// #272: an elevation error during a slew. In the scan of the error only the elevation is disabled and the shared brake is
// closed (no drive holds it); azimuth and derotator stay enabled and get their MC_Stop at the fast-stop dynamics of stMotion
// (bAxisErrorRamp), the hydraulics stay on. After the stop has settled the emergency park parks in place: all axes disabled,
// brake closed, covers closed, hydraulics off, the stop dynamics back at the NC parameters (0.0). Until 0.23.x all three axes
// were disabled in the scan of the error and the brake alone stopped the azimuth.
// #277: the azimuth drive (the NC enable behind the HalfBROT brake gate, fbAxis.Ready in the mock) stays on during the ramp
// although the shared brake is closed (HalfBROT FB_BrakeCloseHold); without the hold the gate dropped it in the next scan.
METHOD PRIVATE Elevation_Error_During_A_Slew_Fast_Stops_The_Healthy_Axes
VAR_INST
	pRig		: POINTER TO FB_MonetRig;	// created with __NEW in this test's turn, freed in the scan it finished in
	rig			: REFERENCE TO FB_MonetRig;
	stCfg		: BROTLib.ST_MotionConfig;
	nStep		: INT;
	nCycles		: UINT;
	sTest		: STRING(80);
	nAz0		: UINT;
	nDr0		: UINT;
	nDisable0	: UINT;
	bSeenError	: BOOL;
	bSawRamp	: BOOL;
	bAzDriveLost	: BOOL;	// #277: a ramp scan with the azimuth wanted enabled but its drive off
END_VAR
TEST('Elevation_Error_During_A_Slew_Fast_Stops_The_Healthy_Axes');
sTest := 'Elevation_Error_During_A_Slew_Fast_Stops_The_Healthy_Axes: ';
IF nStep >= 90 THEN
	RETURN;
END_IF
IF nCur <> 22 THEN	// not this test's turn yet (TEST() above is called in every scan, TcUnit needs that)
	RETURN;
END_IF
IF pRig = 0 THEN
	pRig := __NEW(FB_MonetRig);
	IF pRig = 0 THEN
		AssertTrue(Condition := FALSE, Message := 'no router memory for the rig');
		F_Note(bFailed := TRUE, sText := CONCAT(sTest, 'no router memory for the rig'));
		nStep := 99;
		nCur := nCur + 1;
		TEST_FINISHED();
		RETURN;
	END_IF
	rig REF= pRig^;
END_IF
IF nStep = 0 AND nCycles = 0 THEN
	stCfg.fAzimuthFastStopDeceleration := 10.0;
	stCfg.fAzimuthFastStopJerk := 30.0;
	stCfg.fElevationFastStopDeceleration := 9.0;
	stCfg.fElevationFastStopJerk := 27.0;
	stCfg.fDerotatorFastStopDeceleration := 20.0;
	stCfg.fDerotatorFastStopJerk := 60.0;
	rig.SetMotion(stValue := stCfg);
END_IF
rig.Scan();
nCycles := nCycles + 1;
CASE nStep OF
0:	// wait for the clock, then power on
	IF rig.ClockValid THEN
		rig.fbTel.Init();
		nStep := 10;
		nCycles := 0;
	ELSIF nCycles > 2000 THEN
		AssertTrue(Condition := FALSE, Message := 'the astronomical clock never became valid');
		F_Note(bFailed := TRUE, sText := CONCAT(sTest, 'the astronomical clock never became valid'));
		nStep := 99;
		TEST_FINISHED();
	END_IF
10:	// online: slew
	IF rig.Online THEN
		rig.fbTel.Slew(fAzimuth := 180.0, fAltitude := 45.0);
		nStep := 20;
		nCycles := 0;
	ELSIF nCycles > 1500 THEN
		AssertTrue(Condition := FALSE, Message := 'the mock telescope did not reach READY_STATE 1.0');
		F_Note(bFailed := TRUE, sText := CONCAT(sTest, 'the mock telescope did not reach READY_STATE 1.0'));
		nStep := 99;
		TEST_FINISHED();
	END_IF
20:	// the slew moves all three axes: the elevation reports an error
	IF rig.fbElev.MoveAxis AND rig.fbAzim.MoveAxis AND rig.fbDero.MoveAxis AND nCycles >= 3 THEN
		nAz0 := rig.fbAzim.nStopEdges;
		nDr0 := rig.fbDero.nStopEdges;
		nDisable0 := rig.fbBrakeHyd.nDisableCalls;
		rig.InjectElevationError(16#4550);
		nStep := 30;
		nCycles := 0;
	ELSIF nCycles > 300 THEN
		AssertTrue(Condition := FALSE, Message := 'the slew did not start the axis moves');
		F_Note(bFailed := TRUE, sText := CONCAT(sTest, 'the slew did not start the axis moves'));
		nStep := 99;
		TEST_FINISHED();
	END_IF
30:
	bSawRamp := bSawRamp OR rig.fbTel.bAxisErrorRamp;
	// the drive off while the azimuth still moves or stops (the mock core keeps moving without its enable)
	IF rig.fbTel.bAxisErrorRamp AND rig.fbAzim.bEnable AND NOT rig.fbAzim.fbAxis.Ready AND NOT rig.fbAzim.fbAxis.StandStill THEN
		bAzDriveLost := TRUE;
	END_IF
	IF rig.fbTel.bError AND NOT bSeenError THEN	// the scan that saw the error
		bSeenError := TRUE;
		AssertTrue(Condition := rig.fbTel.bAxisErrorRamp AND rig.fbTel.bStopActive, Message := 'the error starts the ramp (bStop)');
		F_Note(bFailed := NOT (rig.fbTel.bAxisErrorRamp AND rig.fbTel.bStopActive), sText := CONCAT(sTest, 'the error starts the ramp (bStop)'));
		AssertFalse(Condition := rig.fbElev.bEnable, Message := 'the faulty elevation is disabled');
		F_Note(bFailed := (rig.fbElev.bEnable), sText := CONCAT(sTest, 'the faulty elevation is disabled'));
		AssertTrue(Condition := rig.fbAzim.bEnable AND rig.fbDero.bEnable, Message := 'azimuth and derotator stay enabled for their stop');
		F_Note(bFailed := NOT (rig.fbAzim.bEnable AND rig.fbDero.bEnable), sText := CONCAT(sTest, 'azimuth and derotator stay enabled for their stop'));
		AssertFalse(Condition := rig.fbBrakeHyd.BrakeOpen, Message := 'the shared brake is closed at once');
		F_Note(bFailed := (rig.fbBrakeHyd.BrakeOpen), sText := CONCAT(sTest, 'the shared brake is closed at once'));
		AssertTrue(Condition := rig.fbBrakeHyd.nDisableCalls = nDisable0, Message := 'the hydraulics stay on');
		F_Note(bFailed := NOT (rig.fbBrakeHyd.nDisableCalls = nDisable0), sText := CONCAT(sTest, 'the hydraulics stay on'));
		AssertTrue(Condition := rig.fbAzim.fbAxis.StopDeceleration = 10.0 AND rig.fbAzim.fbAxis.StopJerk = 30.0, Message := 'the azimuth stops at its fast-stop dynamics');
		F_Note(bFailed := NOT (rig.fbAzim.fbAxis.StopDeceleration = 10.0 AND rig.fbAzim.fbAxis.StopJerk = 30.0), sText := CONCAT(sTest, 'the azimuth stops at its fast-stop dynamics'));
		AssertTrue(Condition := rig.fbDero.fbAxis.StopDeceleration = 20.0 AND rig.fbDero.fbAxis.StopJerk = 60.0, Message := 'the derotator stops at its fast-stop dynamics');
		F_Note(bFailed := NOT (rig.fbDero.fbAxis.StopDeceleration = 20.0 AND rig.fbDero.fbAxis.StopJerk = 60.0), sText := CONCAT(sTest, 'the derotator stops at its fast-stop dynamics'));
	END_IF
	IF rig.fbTel.bIsParked AND nCycles > 5 THEN
		AssertTrue(Condition := bSawRamp, Message := 'the ramp ran');
		F_Note(bFailed := NOT (bSawRamp), sText := CONCAT(sTest, 'the ramp ran'));
		AssertFalse(Condition := bAzDriveLost, Message := 'the azimuth drive stays on for its stop with the brake closed');
		F_Note(bFailed := bAzDriveLost, sText := CONCAT(sTest, 'the azimuth drive stays on for its stop with the brake closed'));
		AssertTrue(Condition := rig.fbAzim.nStopEdges > nAz0 AND rig.fbDero.nStopEdges > nDr0, Message := 'azimuth and derotator were sent their MC_Stop');
		F_Note(bFailed := NOT (rig.fbAzim.nStopEdges > nAz0 AND rig.fbDero.nStopEdges > nDr0), sText := CONCAT(sTest, 'azimuth and derotator were sent their MC_Stop'));
		AssertTrue(Condition := rig.fbTel.bParkedInPlace AND NOT rig.fbTel.bParkActive AND NOT rig.fbTel.bAxisErrorRamp, Message := 'the park ended in place, the ramp is over');
		F_Note(bFailed := NOT (rig.fbTel.bParkedInPlace AND NOT rig.fbTel.bParkActive AND NOT rig.fbTel.bAxisErrorRamp), sText := CONCAT(sTest, 'the park ended in place, the ramp is over'));
		AssertFalse(Condition := rig.fbElev.bEnable OR rig.fbAzim.bEnable OR rig.fbDero.bEnable, Message := 'all three axes are disabled');
		F_Note(bFailed := (rig.fbElev.bEnable OR rig.fbAzim.bEnable OR rig.fbDero.bEnable), sText := CONCAT(sTest, 'all three axes are disabled'));
		AssertFalse(Condition := rig.fbBrakeHyd.BrakeOpen, Message := 'the brake is closed');
		F_Note(bFailed := (rig.fbBrakeHyd.BrakeOpen), sText := CONCAT(sTest, 'the brake is closed'));
		AssertTrue(Condition := rig.fbCovers.bClosed AND rig.fbBrakeHyd.nDisableCalls > nDisable0, Message := 'covers closed, hydraulics off');
		F_Note(bFailed := NOT (rig.fbCovers.bClosed AND rig.fbBrakeHyd.nDisableCalls > nDisable0), sText := CONCAT(sTest, 'covers closed, hydraulics off'));
		AssertTrue(Condition := rig.fbAzim.fbAxis.StopDeceleration = 0.0 AND rig.fbAzim.fbAxis.StopJerk = 0.0 AND
			rig.fbDero.fbAxis.StopDeceleration = 0.0 AND rig.fbElev.fbAxis.StopDeceleration = 0.0, Message := 'the stop dynamics are back at the NC parameters');
		F_Note(bFailed := NOT (rig.fbAzim.fbAxis.StopDeceleration = 0.0 AND rig.fbAzim.fbAxis.StopJerk = 0.0 AND
			rig.fbDero.fbAxis.StopDeceleration = 0.0 AND rig.fbElev.fbAxis.StopDeceleration = 0.0), sText := CONCAT(sTest, 'the stop dynamics are back at the NC parameters'));
		AssertTrue(Condition := rig.fbTel.bError AND rig.fbTel.ReadyState = -1.0, Message := 'the error stays, READY_STATE -1.0');
		F_Note(bFailed := NOT (rig.fbTel.bError AND rig.fbTel.ReadyState = -1.0), sText := CONCAT(sTest, 'the error stays, READY_STATE -1.0'));
		nStep := 99;
		TEST_FINISHED();
	ELSIF nCycles > 1000 THEN
		AssertTrue(Condition := FALSE, Message := 'the telescope did not park after the ramp');
		F_Note(bFailed := TRUE, sText := CONCAT(sTest, 'the telescope did not park after the ramp'));
		nStep := 99;
		TEST_FINISHED();
	END_IF
END_CASE
IF nStep >= 90 AND pRig <> 0 THEN	// finished in this scan: free the rig, the next test starts in the next scan
	__DELETE(pRig);
	pRig := 0;
	nCur := nCur + 1;
END_IF
END_METHOD

// #272: an azimuth error during a slew. The faulty azimuth has no drive, so the shared brake is closed in the scan of the error
// (until 0.23.x the emergency park closed it in that scan; the park now waits behind the ramp) and held closed: the enabled
// elevation requests the opening in every scan. Elevation and derotator stay enabled and get their MC_Stop; then the park parks
// in place. #277: the elevation drive stays on for its stop although the brake is closed (HalfBROT FB_BrakeCloseHold).
METHOD PRIVATE Azimuth_Error_During_A_Slew_Closes_The_Brake_At_Once
VAR_INST
	pRig		: POINTER TO FB_MonetRig;	// created with __NEW in this test's turn, freed in the scan it finished in
	rig			: REFERENCE TO FB_MonetRig;
	nStep		: INT;
	nCycles		: UINT;
	sTest		: STRING(80);
	nEl0		: UINT;
	nDisable0	: UINT;
	bSeenError	: BOOL;
	bReopened	: BOOL;	// the brake was open again in a later scan of the ramp (the enabled elevation requests the opening in every scan)
	bElDriveLost	: BOOL;	// #277: a ramp scan with the elevation wanted enabled but its drive off while it still moves
END_VAR
TEST('Azimuth_Error_During_A_Slew_Closes_The_Brake_At_Once');
sTest := 'Azimuth_Error_During_A_Slew_Closes_The_Brake_At_Once: ';
IF nStep >= 90 THEN
	RETURN;
END_IF
IF nCur <> 23 THEN	// not this test's turn yet (TEST() above is called in every scan, TcUnit needs that)
	RETURN;
END_IF
IF pRig = 0 THEN
	pRig := __NEW(FB_MonetRig);
	IF pRig = 0 THEN
		AssertTrue(Condition := FALSE, Message := 'no router memory for the rig');
		F_Note(bFailed := TRUE, sText := CONCAT(sTest, 'no router memory for the rig'));
		nStep := 99;
		nCur := nCur + 1;
		TEST_FINISHED();
		RETURN;
	END_IF
	rig REF= pRig^;
END_IF
rig.Scan();
nCycles := nCycles + 1;
CASE nStep OF
0:	// wait for the clock, then power on
	IF rig.ClockValid THEN
		rig.fbTel.Init();
		nStep := 10;
		nCycles := 0;
	ELSIF nCycles > 2000 THEN
		AssertTrue(Condition := FALSE, Message := 'the astronomical clock never became valid');
		F_Note(bFailed := TRUE, sText := CONCAT(sTest, 'the astronomical clock never became valid'));
		nStep := 99;
		TEST_FINISHED();
	END_IF
10:	// online: slew
	IF rig.Online THEN
		rig.fbTel.Slew(fAzimuth := 180.0, fAltitude := 45.0);
		nStep := 20;
		nCycles := 0;
	ELSIF nCycles > 1500 THEN
		AssertTrue(Condition := FALSE, Message := 'the mock telescope did not reach READY_STATE 1.0');
		F_Note(bFailed := TRUE, sText := CONCAT(sTest, 'the mock telescope did not reach READY_STATE 1.0'));
		nStep := 99;
		TEST_FINISHED();
	END_IF
20:	// the slew moves all three axes: the azimuth reports an error
	IF rig.fbElev.MoveAxis AND rig.fbAzim.MoveAxis AND rig.fbDero.MoveAxis AND nCycles >= 3 THEN
		nEl0 := rig.fbElev.nStopEdges;
		nDisable0 := rig.fbBrakeHyd.nDisableCalls;
		rig.InjectAzimuthError(16#4550);
		nStep := 30;
		nCycles := 0;
	ELSIF nCycles > 300 THEN
		AssertTrue(Condition := FALSE, Message := 'the slew did not start the axis moves');
		F_Note(bFailed := TRUE, sText := CONCAT(sTest, 'the slew did not start the axis moves'));
		nStep := 99;
		TEST_FINISHED();
	END_IF
30:
	IF rig.fbTel.bAxisErrorRamp AND rig.fbElev.bEnable AND NOT rig.fbElev.fbAxis.Ready AND NOT rig.fbElev.fbAxis.StandStill THEN
		bElDriveLost := TRUE;
	END_IF
	IF rig.fbTel.bError AND NOT bSeenError THEN	// the scan that saw the error
		bSeenError := TRUE;
		AssertTrue(Condition := rig.fbTel.bAxisErrorRamp, Message := 'the error starts the ramp');
		F_Note(bFailed := NOT (rig.fbTel.bAxisErrorRamp), sText := CONCAT(sTest, 'the error starts the ramp'));
		AssertFalse(Condition := rig.fbAzim.bEnable, Message := 'the faulty azimuth is disabled');
		F_Note(bFailed := (rig.fbAzim.bEnable), sText := CONCAT(sTest, 'the faulty azimuth is disabled'));
		AssertTrue(Condition := rig.fbElev.bEnable AND rig.fbDero.bEnable, Message := 'elevation and derotator stay enabled for their stop');
		F_Note(bFailed := NOT (rig.fbElev.bEnable AND rig.fbDero.bEnable), sText := CONCAT(sTest, 'elevation and derotator stay enabled for their stop'));
		AssertFalse(Condition := rig.fbBrakeHyd.BrakeOpen, Message := 'the shared brake is closed at once');
		F_Note(bFailed := (rig.fbBrakeHyd.BrakeOpen), sText := CONCAT(sTest, 'the shared brake is closed at once'));
		AssertTrue(Condition := rig.fbBrakeHyd.nDisableCalls = nDisable0, Message := 'the hydraulics stay on');
		F_Note(bFailed := NOT (rig.fbBrakeHyd.nDisableCalls = nDisable0), sText := CONCAT(sTest, 'the hydraulics stay on'));
	ELSIF bSeenError AND rig.fbBrakeHyd.BrakeOpen THEN
		bReopened := TRUE;
	END_IF
	IF rig.fbTel.bIsParked AND nCycles > 5 THEN
		AssertFalse(Condition := bReopened, Message := 'the brake stays closed after the error');
		F_Note(bFailed := bReopened, sText := CONCAT(sTest, 'the brake stays closed after the error'));
		AssertFalse(Condition := bElDriveLost, Message := 'the elevation drive stays on for its stop with the brake closed');
		F_Note(bFailed := bElDriveLost, sText := CONCAT(sTest, 'the elevation drive stays on for its stop with the brake closed'));
		AssertTrue(Condition := bSeenError AND rig.fbElev.nStopEdges > nEl0, Message := 'the elevation was sent its MC_Stop');
		F_Note(bFailed := NOT (bSeenError AND rig.fbElev.nStopEdges > nEl0), sText := CONCAT(sTest, 'the elevation was sent its MC_Stop'));
		AssertTrue(Condition := rig.fbTel.bParkedInPlace AND NOT rig.fbTel.bParkActive, Message := 'the park ended in place');
		F_Note(bFailed := NOT (rig.fbTel.bParkedInPlace AND NOT rig.fbTel.bParkActive), sText := CONCAT(sTest, 'the park ended in place'));
		AssertFalse(Condition := rig.fbElev.bEnable OR rig.fbAzim.bEnable OR rig.fbDero.bEnable, Message := 'all three axes are disabled');
		F_Note(bFailed := (rig.fbElev.bEnable OR rig.fbAzim.bEnable OR rig.fbDero.bEnable), sText := CONCAT(sTest, 'all three axes are disabled'));
		AssertTrue(Condition := rig.fbCovers.bClosed AND rig.fbBrakeHyd.nDisableCalls > nDisable0, Message := 'covers closed, hydraulics off');
		F_Note(bFailed := NOT (rig.fbCovers.bClosed AND rig.fbBrakeHyd.nDisableCalls > nDisable0), sText := CONCAT(sTest, 'covers closed, hydraulics off'));
		nStep := 99;
		TEST_FINISHED();
	ELSIF nCycles > 1000 THEN
		AssertTrue(Condition := FALSE, Message := 'the telescope did not park after the ramp');
		F_Note(bFailed := TRUE, sText := CONCAT(sTest, 'the telescope did not park after the ramp'));
		nStep := 99;
		TEST_FINISHED();
	END_IF
END_CASE
IF nStep >= 90 AND pRig <> 0 THEN	// finished in this scan: free the rig, the next test starts in the next scan
	__DELETE(pRig);
	pRig := 0;
	nCur := nCur + 1;
END_IF
END_METHOD

// #272: a derotator error alone during a slew. The derotator is not on the hydraulic brake: the brake stays open and the
// hydraulics on while elevation and azimuth stop with their drives; the park in place closes the brake at rest.
METHOD PRIVATE Derotator_Error_During_A_Slew_Keeps_The_Brake_Open_For_The_Ramp
VAR_INST
	pRig		: POINTER TO FB_MonetRig;	// created with __NEW in this test's turn, freed in the scan it finished in
	rig			: REFERENCE TO FB_MonetRig;
	nStep		: INT;
	nCycles		: UINT;
	sTest		: STRING(80);
	nEl0		: UINT;
	nAz0		: UINT;
	nDisable0	: UINT;
	bSeenError	: BOOL;
END_VAR
TEST('Derotator_Error_During_A_Slew_Keeps_The_Brake_Open_For_The_Ramp');
sTest := 'Derotator_Error_During_A_Slew_Keeps_The_Brake_Open_For_The_Ramp: ';
IF nStep >= 90 THEN
	RETURN;
END_IF
IF nCur <> 24 THEN	// not this test's turn yet (TEST() above is called in every scan, TcUnit needs that)
	RETURN;
END_IF
IF pRig = 0 THEN
	pRig := __NEW(FB_MonetRig);
	IF pRig = 0 THEN
		AssertTrue(Condition := FALSE, Message := 'no router memory for the rig');
		F_Note(bFailed := TRUE, sText := CONCAT(sTest, 'no router memory for the rig'));
		nStep := 99;
		nCur := nCur + 1;
		TEST_FINISHED();
		RETURN;
	END_IF
	rig REF= pRig^;
END_IF
rig.Scan();
nCycles := nCycles + 1;
CASE nStep OF
0:	// wait for the clock, then power on
	IF rig.ClockValid THEN
		rig.fbTel.Init();
		nStep := 10;
		nCycles := 0;
	ELSIF nCycles > 2000 THEN
		AssertTrue(Condition := FALSE, Message := 'the astronomical clock never became valid');
		F_Note(bFailed := TRUE, sText := CONCAT(sTest, 'the astronomical clock never became valid'));
		nStep := 99;
		TEST_FINISHED();
	END_IF
10:	// online: slew
	IF rig.Online THEN
		rig.fbTel.Slew(fAzimuth := 180.0, fAltitude := 45.0);
		nStep := 20;
		nCycles := 0;
	ELSIF nCycles > 1500 THEN
		AssertTrue(Condition := FALSE, Message := 'the mock telescope did not reach READY_STATE 1.0');
		F_Note(bFailed := TRUE, sText := CONCAT(sTest, 'the mock telescope did not reach READY_STATE 1.0'));
		nStep := 99;
		TEST_FINISHED();
	END_IF
20:	// the slew moves all three axes: the derotator reports an error
	IF rig.fbElev.MoveAxis AND rig.fbAzim.MoveAxis AND rig.fbDero.MoveAxis AND nCycles >= 3 THEN
		nEl0 := rig.fbElev.nStopEdges;
		nAz0 := rig.fbAzim.nStopEdges;
		nDisable0 := rig.fbBrakeHyd.nDisableCalls;
		rig.InjectDerotatorError(16#4550);
		nStep := 30;
		nCycles := 0;
	ELSIF nCycles > 300 THEN
		AssertTrue(Condition := FALSE, Message := 'the slew did not start the axis moves');
		F_Note(bFailed := TRUE, sText := CONCAT(sTest, 'the slew did not start the axis moves'));
		nStep := 99;
		TEST_FINISHED();
	END_IF
30:
	IF rig.fbTel.bError AND NOT bSeenError THEN	// the scan that saw the error
		bSeenError := TRUE;
		AssertTrue(Condition := rig.fbTel.bAxisErrorRamp, Message := 'the error starts the ramp');
		F_Note(bFailed := NOT (rig.fbTel.bAxisErrorRamp), sText := CONCAT(sTest, 'the error starts the ramp'));
		AssertFalse(Condition := rig.fbDero.bEnable, Message := 'the faulty derotator is disabled');
		F_Note(bFailed := (rig.fbDero.bEnable), sText := CONCAT(sTest, 'the faulty derotator is disabled'));
		AssertTrue(Condition := rig.fbElev.bEnable AND rig.fbAzim.bEnable, Message := 'elevation and azimuth stay enabled for their stop');
		F_Note(bFailed := NOT (rig.fbElev.bEnable AND rig.fbAzim.bEnable), sText := CONCAT(sTest, 'elevation and azimuth stay enabled for their stop'));
		AssertTrue(Condition := rig.fbBrakeHyd.BrakeOpen AND rig.fbBrakeHyd.nDisableCalls = nDisable0, Message := 'the brake stays open and the hydraulics on');
		F_Note(bFailed := NOT (rig.fbBrakeHyd.BrakeOpen AND rig.fbBrakeHyd.nDisableCalls = nDisable0), sText := CONCAT(sTest, 'the brake stays open and the hydraulics on'));
	END_IF
	IF rig.fbTel.bIsParked AND nCycles > 5 THEN
		AssertTrue(Condition := bSeenError AND rig.fbElev.nStopEdges > nEl0 AND rig.fbAzim.nStopEdges > nAz0, Message := 'elevation and azimuth were sent their MC_Stop');
		F_Note(bFailed := NOT (bSeenError AND rig.fbElev.nStopEdges > nEl0 AND rig.fbAzim.nStopEdges > nAz0), sText := CONCAT(sTest, 'elevation and azimuth were sent their MC_Stop'));
		AssertTrue(Condition := rig.fbTel.bParkedInPlace AND NOT rig.fbTel.bParkActive, Message := 'the park ended in place');
		F_Note(bFailed := NOT (rig.fbTel.bParkedInPlace AND NOT rig.fbTel.bParkActive), sText := CONCAT(sTest, 'the park ended in place'));
		AssertFalse(Condition := rig.fbElev.bEnable OR rig.fbAzim.bEnable OR rig.fbDero.bEnable, Message := 'all three axes are disabled');
		F_Note(bFailed := (rig.fbElev.bEnable OR rig.fbAzim.bEnable OR rig.fbDero.bEnable), sText := CONCAT(sTest, 'all three axes are disabled'));
		AssertFalse(Condition := rig.fbBrakeHyd.BrakeOpen, Message := 'the brake is closed at rest');
		F_Note(bFailed := (rig.fbBrakeHyd.BrakeOpen), sText := CONCAT(sTest, 'the brake is closed at rest'));
		AssertTrue(Condition := rig.fbCovers.bClosed AND rig.fbBrakeHyd.nDisableCalls > nDisable0, Message := 'covers closed, hydraulics off');
		F_Note(bFailed := NOT (rig.fbCovers.bClosed AND rig.fbBrakeHyd.nDisableCalls > nDisable0), sText := CONCAT(sTest, 'covers closed, hydraulics off'));
		nStep := 99;
		TEST_FINISHED();
	ELSIF nCycles > 1000 THEN
		AssertTrue(Condition := FALSE, Message := 'the telescope did not park after the ramp');
		F_Note(bFailed := TRUE, sText := CONCAT(sTest, 'the telescope did not park after the ramp'));
		nStep := 99;
		TEST_FINISHED();
	END_IF
END_CASE
IF nStep >= 90 AND pRig <> 0 THEN	// finished in this scan: free the rig, the next test starts in the next scan
	__DELETE(pRig);
	pRig := 0;
	nCur := nCur + 1;
END_IF
END_METHOD

// #272: a further axis error during the ramp of an axis error ends the ramp: the error branch disables all three axes, as
// before 0.24. The stops are made slow (SetStopScans 200) so that the ramp is still running when the azimuth faults.
METHOD PRIVATE Second_Axis_Error_During_The_Ramp_Disables_All_Axes
VAR_INST
	pRig		: POINTER TO FB_MonetRig;	// created with __NEW in this test's turn, freed in the scan it finished in
	rig			: REFERENCE TO FB_MonetRig;
	nStep		: INT;
	nCycles		: UINT;
	sTest		: STRING(80);
END_VAR
TEST('Second_Axis_Error_During_The_Ramp_Disables_All_Axes');
sTest := 'Second_Axis_Error_During_The_Ramp_Disables_All_Axes: ';
IF nStep >= 90 THEN
	RETURN;
END_IF
IF nCur <> 25 THEN	// not this test's turn yet (TEST() above is called in every scan, TcUnit needs that)
	RETURN;
END_IF
IF pRig = 0 THEN
	pRig := __NEW(FB_MonetRig);
	IF pRig = 0 THEN
		AssertTrue(Condition := FALSE, Message := 'no router memory for the rig');
		F_Note(bFailed := TRUE, sText := CONCAT(sTest, 'no router memory for the rig'));
		nStep := 99;
		nCur := nCur + 1;
		TEST_FINISHED();
		RETURN;
	END_IF
	rig REF= pRig^;
END_IF
rig.Scan();
nCycles := nCycles + 1;
CASE nStep OF
0:	// wait for the clock, then power on
	IF rig.ClockValid THEN
		rig.fbTel.Init();
		nStep := 10;
		nCycles := 0;
	ELSIF nCycles > 2000 THEN
		AssertTrue(Condition := FALSE, Message := 'the astronomical clock never became valid');
		F_Note(bFailed := TRUE, sText := CONCAT(sTest, 'the astronomical clock never became valid'));
		nStep := 99;
		TEST_FINISHED();
	END_IF
10:	// online: slew with slow stops
	IF rig.Online THEN
		rig.SetStopScans(nScans := 200);
		rig.fbTel.Slew(fAzimuth := 180.0, fAltitude := 45.0);
		nStep := 20;
		nCycles := 0;
	ELSIF nCycles > 1500 THEN
		AssertTrue(Condition := FALSE, Message := 'the mock telescope did not reach READY_STATE 1.0');
		F_Note(bFailed := TRUE, sText := CONCAT(sTest, 'the mock telescope did not reach READY_STATE 1.0'));
		nStep := 99;
		TEST_FINISHED();
	END_IF
20:	// the slew moves all three axes: the elevation reports an error
	IF rig.fbElev.MoveAxis AND rig.fbAzim.MoveAxis AND rig.fbDero.MoveAxis AND nCycles >= 3 THEN
		rig.InjectElevationError(16#4550);
		nStep := 30;
		nCycles := 0;
	ELSIF nCycles > 300 THEN
		AssertTrue(Condition := FALSE, Message := 'the slew did not start the axis moves');
		F_Note(bFailed := TRUE, sText := CONCAT(sTest, 'the slew did not start the axis moves'));
		nStep := 99;
		TEST_FINISHED();
	END_IF
30:	// the ramp runs: the azimuth faults too
	IF nCycles >= 5 THEN
		AssertTrue(Condition := rig.fbTel.bAxisErrorRamp AND rig.fbAzim.bEnable, Message := 'the ramp of the elevation error runs');
		F_Note(bFailed := NOT (rig.fbTel.bAxisErrorRamp AND rig.fbAzim.bEnable), sText := CONCAT(sTest, 'the ramp of the elevation error runs'));
		rig.InjectAzimuthError(16#4550);
		nStep := 40;
		nCycles := 0;
	END_IF
40:	// within two scans the ramp is over and all axes are disabled
	IF nCycles >= 2 THEN
		AssertFalse(Condition := rig.fbTel.bAxisErrorRamp, Message := 'the second error ends the ramp');
		F_Note(bFailed := (rig.fbTel.bAxisErrorRamp), sText := CONCAT(sTest, 'the second error ends the ramp'));
		AssertFalse(Condition := rig.fbElev.bEnable OR rig.fbAzim.bEnable OR rig.fbDero.bEnable, Message := 'all three axes are disabled');
		F_Note(bFailed := (rig.fbElev.bEnable OR rig.fbAzim.bEnable OR rig.fbDero.bEnable), sText := CONCAT(sTest, 'all three axes are disabled'));
		nStep := 99;
		TEST_FINISHED();
	END_IF
END_CASE
IF nStep >= 90 AND pRig <> 0 THEN	// finished in this scan: free the rig, the next test starts in the next scan
	__DELETE(pRig);
	pRig := 0;
	nCur := nCur + 1;
END_IF
END_METHOD

// #277, the order of MONET/N run B (2026-11-13, an ADS write ElevationControl.bEnable := FALSE during a slew): the elevation
// is disabled first, HalfBROT closes the shared brake on the falling edge of its enable, and the elevation error is seen one scan
// later, with the brake already closed. The azimuth keeps its drive through the closing (HalfBROT FB_BrakeCloseHold), so the ramp
// still starts (until 0.24.0 it needed the brake open on the error edge, and the azimuth was disabled and braked from slew speed)
// and the azimuth gets its MC_Stop with the drive on; then the park parks in place.
METHOD PRIVATE Elevation_Disabled_Before_Its_Error_Still_Fast_Stops_The_Azimuth
VAR_INST
	pRig		: POINTER TO FB_MonetRig;	// created with __NEW in this test's turn, freed in the scan it finished in
	rig			: REFERENCE TO FB_MonetRig;
	nStep		: INT;
	nCycles		: UINT;
	sTest		: STRING(80);
	nAz0		: UINT;
	bSawRamp	: BOOL;
	bAzDriveLost	: BOOL;	// a scan with the azimuth wanted enabled but its drive off while it still moves (before the park disables it)
END_VAR
TEST('Elevation_Disabled_Before_Its_Error_Still_Fast_Stops_The_Azimuth');
sTest := 'Elevation_Disabled_Before_Its_Error_Still_Fast_Stops_The_Azimuth: ';
IF nStep >= 90 THEN
	RETURN;
END_IF
IF nCur <> 26 THEN	// not this test's turn yet (TEST() above is called in every scan, TcUnit needs that)
	RETURN;
END_IF
IF pRig = 0 THEN
	pRig := __NEW(FB_MonetRig);
	IF pRig = 0 THEN
		AssertTrue(Condition := FALSE, Message := 'no router memory for the rig');
		F_Note(bFailed := TRUE, sText := CONCAT(sTest, 'no router memory for the rig'));
		nStep := 99;
		nCur := nCur + 1;
		TEST_FINISHED();
		RETURN;
	END_IF
	rig REF= pRig^;
END_IF
rig.Scan();
nCycles := nCycles + 1;
IF nStep >= 25 AND nStep < 90 THEN
	bSawRamp := bSawRamp OR rig.fbTel.bAxisErrorRamp;
	IF rig.fbAzim.bEnable AND NOT rig.fbAzim.fbAxis.Ready AND NOT rig.fbAzim.fbAxis.StandStill THEN
		bAzDriveLost := TRUE;
	END_IF
END_IF
CASE nStep OF
0:	// wait for the clock, then power on
	IF rig.ClockValid THEN
		rig.fbTel.Init();
		nStep := 10;
		nCycles := 0;
	ELSIF nCycles > 2000 THEN
		AssertTrue(Condition := FALSE, Message := 'the astronomical clock never became valid');
		F_Note(bFailed := TRUE, sText := CONCAT(sTest, 'the astronomical clock never became valid'));
		nStep := 99;
		TEST_FINISHED();
	END_IF
10:	// online: slew
	IF rig.Online THEN
		rig.fbTel.Slew(fAzimuth := 180.0, fAltitude := 45.0);
		nStep := 20;
		nCycles := 0;
	ELSIF nCycles > 1500 THEN
		AssertTrue(Condition := FALSE, Message := 'the mock telescope did not reach READY_STATE 1.0');
		F_Note(bFailed := TRUE, sText := CONCAT(sTest, 'the mock telescope did not reach READY_STATE 1.0'));
		nStep := 99;
		TEST_FINISHED();
	END_IF
20:	// the slew moves all three axes: the elevation enable drops (the ADS write of run B)
	IF rig.fbElev.MoveAxis AND rig.fbAzim.MoveAxis AND rig.fbDero.MoveAxis AND nCycles >= 3 THEN
		nAz0 := rig.fbAzim.nStopEdges;
		rig.DisableElevation();
		nStep := 25;
		nCycles := 0;
	ELSIF nCycles > 300 THEN
		AssertTrue(Condition := FALSE, Message := 'the slew did not start the axis moves');
		F_Note(bFailed := TRUE, sText := CONCAT(sTest, 'the slew did not start the axis moves'));
		nStep := 99;
		TEST_FINISHED();
	END_IF
25:	// one scan later: the brake is closed, the azimuth still has its drive; now the elevation reports its error
	AssertFalse(Condition := rig.fbBrakeHyd.BrakeOpen, Message := 'the falling enable closed the brake');
	F_Note(bFailed := rig.fbBrakeHyd.BrakeOpen, sText := CONCAT(sTest, 'the falling enable closed the brake'));
	AssertTrue(Condition := rig.fbAzim.fbAxis.Ready, Message := 'the moving azimuth keeps its drive through the closing');
	F_Note(bFailed := NOT rig.fbAzim.fbAxis.Ready, sText := CONCAT(sTest, 'the moving azimuth keeps its drive through the closing'));
	rig.InjectElevationError(16#4260);
	nStep := 30;
	nCycles := 0;
30:
	IF rig.fbTel.bIsParked AND nCycles > 5 THEN
		AssertTrue(Condition := bSawRamp, Message := 'the ramp ran although the brake was closed on the error edge');
		F_Note(bFailed := NOT bSawRamp, sText := CONCAT(sTest, 'the ramp ran although the brake was closed on the error edge'));
		AssertTrue(Condition := rig.fbAzim.nStopEdges > nAz0, Message := 'the azimuth was sent its MC_Stop');
		F_Note(bFailed := NOT (rig.fbAzim.nStopEdges > nAz0), sText := CONCAT(sTest, 'the azimuth was sent its MC_Stop'));
		AssertFalse(Condition := bAzDriveLost, Message := 'the azimuth drive stays on until it stands');
		F_Note(bFailed := bAzDriveLost, sText := CONCAT(sTest, 'the azimuth drive stays on until it stands'));
		AssertTrue(Condition := rig.fbTel.bParkedInPlace AND NOT rig.fbTel.bParkActive, Message := 'the park ended in place');
		F_Note(bFailed := NOT (rig.fbTel.bParkedInPlace AND NOT rig.fbTel.bParkActive), sText := CONCAT(sTest, 'the park ended in place'));
		AssertFalse(Condition := rig.fbElev.bEnable OR rig.fbAzim.bEnable OR rig.fbDero.bEnable, Message := 'all three axes are disabled');
		F_Note(bFailed := (rig.fbElev.bEnable OR rig.fbAzim.bEnable OR rig.fbDero.bEnable), sText := CONCAT(sTest, 'all three axes are disabled'));
		AssertFalse(Condition := rig.fbBrakeHyd.BrakeOpen, Message := 'the brake is closed');
		F_Note(bFailed := (rig.fbBrakeHyd.BrakeOpen), sText := CONCAT(sTest, 'the brake is closed'));
		nStep := 99;
		TEST_FINISHED();
	ELSIF nCycles > 1000 THEN
		AssertTrue(Condition := FALSE, Message := 'the telescope did not park after the ramp');
		F_Note(bFailed := TRUE, sText := CONCAT(sTest, 'the telescope did not park after the ramp'));
		nStep := 99;
		TEST_FINISHED();
	END_IF
END_CASE
IF nStep >= 90 AND pRig <> 0 THEN	// finished in this scan: free the rig, the next test starts in the next scan
	__DELETE(pRig);
	pRig := 0;
	nCur := nCur + 1;
END_IF
END_METHOD

END_FUNCTION_BLOCK

(* stored: Version 1.1.0.1, ProductVersion 3.1.4024.15
   POU MonetErrorPark_Tests: Id {589804fc-1ef2-48cc-9923-fb6abcd872c3}, SpecialFunc None
   Method Elevation_Error_Starts_The_Emergency_Park: Id {6190de19-41df-490b-93bf-4ae2a295f3a2}
   Method Focus_Error_At_Standstill_Parks_At_The_Park_Position: Id {01032966-7411-4af2-a4d4-6b95b60bd9ac}
   Method Error_On_A_Parked_Telescope_Does_Not_Park_Again: Id {e378877b-adb5-4ca0-af7e-8f895f4ccb2a}
   Method Error_During_Estop_Does_Not_Park: Id {68bf4dbd-82a2-4cd3-ab08-78009e7319a9}
   Method First_PowerOn_AzEl_Error_Is_Exempt_From_The_Park: Id {b161a719-4601-485d-bf30-7cc1d9352e31}
   Method Persisting_Error_Does_Not_Start_A_Second_Park: Id {bccaf610-8410-4c63-88c9-7ae833230e4e}
   Method Power_Failure_At_Standstill_Parks_In_Place_And_Recovers: Id {03d8a622-feb0-4c12-acf2-b4166da20358}
   Method Power_Failure_On_A_Parked_Telescope_Does_Not_Park: Id {be6ce1f6-02e4-4999-ac37-896b59fe2c10}
   Method Hydraulics_Error_On_A_Parked_Telescope_Does_Not_Park: Id {46d579f6-fa1a-4401-a192-f55339d8302e}
   Method Hydraulics_Error_During_Estop_Does_Not_Park: Id {f1554025-9250-4236-b5a5-c6dc739a8ade}
   Method Hydraulics_Error_Park_Recovers_With_Hydraulics_Reset_And_Reset: Id {aa897218-649e-4f97-902a-7d1fe57600a9}
   Method Cover_Error_Park_Recovers_With_Cover_Reset_And_Reset: Id {1aed1f73-4b16-497e-b0a9-80d683867dc4}
   Method Cover_Error_During_Estop_Does_Not_Park: Id {44fb406b-6817-4fcc-830a-795da88a3e6b}
   Method Focus_Error_While_Tracking_Ramps_Then_Parks_At_The_Park_Position: Id {df2e8595-d308-4712-bc6a-f74d383712cd}
   Method Focus_Error_With_An_Axis_Error_Parks_In_Place: Id {f2528670-bf25-467f-ab22-a862eb2d87ea}
   Method Axis_Error_During_The_Focus_Error_Park_Parks_In_Place: Id {f366f26e-855b-4284-9ac6-0481c3eff100}
   Method Stuck_Focus_Does_Not_Hold_The_Focus_Error_Park: Id {ec8b9bca-0bc5-47ed-8a5f-4d900094c09a}
   Method Focus_Error_Park_Recovers_With_Reset_And_Power_On: Id {c890cb45-3f8c-4307-b056-83bf2d5413d9}
   Method Estop_During_Cover_Opening_Stops_The_Covers: Id {a69c945c-64a6-4178-860d-73d39306efcc}
   Method Safety_Error_During_Cover_Opening_Stops_The_Covers: Id {d061df57-c3bc-4c14-b2fb-547df41e2014}
   Method Estop_During_Cover_Closing_Stops_The_Covers: Id {3384dc23-449b-41e7-922b-23cd80459489}
   Method Elevation_Error_During_A_Slew_Fast_Stops_The_Healthy_Axes: Id {19cc2cd3-08a1-4701-8de2-464a0c4f9f7a}
   Method Azimuth_Error_During_A_Slew_Closes_The_Brake_At_Once: Id {005ca04b-8d1d-4d6a-b6aa-bc9fc742bd70}
   Method Derotator_Error_During_A_Slew_Keeps_The_Brake_Open_For_The_Ramp: Id {5322b58c-fd98-49c2-9f7f-9ddec7abfca1}
   Method Second_Axis_Error_During_The_Ramp_Disables_All_Axes: Id {d4229a9e-6bfd-4a1f-9d05-46ac6626f542}
   Method Elevation_Disabled_Before_Its_Error_Still_Fast_Stops_The_Azimuth: Id {39fc59e4-6e09-428a-8d5c-470c5ef9902d} *)
